(* IEC 61131-3 sources: TwinAxisLab/openplc/cobot-6dof-smart-demo, 8 files *)

(* ---- cobot_6dof_iot_condition_monitoring.st ---- *)
VAR
  Command AT %QW90 : UINT := 0;
  Status AT %QW91 : UINT := 0;
  ActiveStep AT %QW92 : UINT := 0;
  ElapsedMsOut AT %QW93 : UINT := 0;
  AlarmCode AT %QW94 : UINT := 0;
  ConditionState AT %QW95 : UINT := 3;
  SpeedPermille AT %QW96 : UINT := 0;
  ProgramSignature AT %QW97 : UINT := 2101;
  J1Raw AT %QW100 : INT := 0;
  J2Raw AT %QW101 : INT := 0;
  J3Raw AT %QW102 : INT := 0;
  J4Raw AT %QW103 : INT := 0;
  J5Raw AT %QW104 : INT := 0;
  J6Raw AT %QW105 : INT := 0;
  TemperatureCx100 AT %QW120 : INT := 0;
  HumidityRHx100 AT %QW121 : UINT := 0;
  GyroDpsx100 AT %QW122 : UINT := 0;
  SensorAgeMs AT %QW123 : UINT := 65535;
  SensorValid AT %QW124 : UINT := 0;
  SensorSequence AT %QW125 : UINT := 0;
  SensorQualityBits AT %QW126 : UINT := 0;
  SensorPolicy AT %QW127 : UINT := 0;
  CycleTimer : TON;
  MotionIdleTimer : TON;
  TimerEnabled : BOOL := FALSE;
  ResetTimer : BOOL := TRUE;
  ElapsedMs : DINT := 0;
  SegmentStartMs : DINT := 0;
  SegmentDurationMs : DINT := 1;
  P : REAL := 0.0;
  MotionScale : REAL := 1.0;
  TemperatureC : REAL := 0.0;
  HumidityRH : REAL := 0.0;
  GyroDps : REAL := 0.0;
  J1Deg : REAL := 0.0;
  J2Deg : REAL := -35.0;
  J3Deg : REAL := 75.0;
  J4Deg : REAL := 50.0;
  J5Deg : REAL := 0.0;
  J6Deg : REAL := 0.0;
  TargetJ1 : REAL := 0.0;
  TargetJ2 : REAL := -35.0;
  TargetJ3 : REAL := 75.0;
  TargetJ4 : REAL := 50.0;
  TargetJ5 : REAL := 0.0;
  TargetJ6 : REAL := 0.0;
  SegmentStartJ1 : REAL := 0.0;
  SegmentStartJ2 : REAL := -35.0;
  SegmentStartJ3 : REAL := 75.0;
  SegmentStartJ4 : REAL := 50.0;
  SegmentStartJ5 : REAL := 0.0;
  SegmentStartJ6 : REAL := 0.0;
  PreviousStep : UINT := 0;
  PreviousP : REAL := 0.0;
  ProgressDelta : REAL := 0.0;
  MotionPresent : BOOL := FALSE;
  DegToRadScaled : REAL := 174.5329;
END_VAR

ProgramSignature := 2101;

TemperatureC := INT_TO_REAL(TemperatureCx100) / 100.0;
HumidityRH := UINT_TO_REAL(HumidityRHx100) / 100.0;
GyroDps := UINT_TO_REAL(GyroDpsx100) / 100.0;
MotionPresent := GyroDps >= 3.0;
MotionIdleTimer(IN := NOT MotionPresent, PT := T#2s);

ConditionState := 0;
AlarmCode := 0;
MotionScale := 1.0;
SpeedPermille := 1000;

IF (SensorValid = 0) OR ((SensorQualityBits AND 1) = 0) OR (SensorAgeMs > 2500) THEN
  ConditionState := 3;
  AlarmCode := 4;
  MotionScale := 0.0;
  SpeedPermille := 0;
ELSIF ((SensorPolicy = 0) OR (SensorPolicy = 1)) AND ((SensorQualityBits AND 16) = 0) THEN
  ConditionState := 3;
  AlarmCode := 6;
  MotionScale := 0.0;
  SpeedPermille := 0;
ELSIF (TemperatureC >= 55.0) OR (HumidityRH >= 85.0) OR (GyroDps >= 220.0) THEN
  ConditionState := 2;
  MotionScale := 0.0;
  SpeedPermille := 0;
  IF TemperatureC >= 55.0 THEN
    AlarmCode := 1;
  ELSIF HumidityRH >= 85.0 THEN
    AlarmCode := 2;
  ELSE
    AlarmCode := 3;
  END_IF;
ELSIF (TemperatureC >= 45.0) OR (HumidityRH >= 75.0) OR (GyroDps >= 120.0) THEN
  ConditionState := 1;
  MotionScale := 0.55;
  SpeedPermille := 550;
ELSIF (SensorPolicy = 0) AND (NOT MotionPresent) AND (NOT MotionIdleTimer.Q) THEN
  ConditionState := 2;
  AlarmCode := 5;
  MotionScale := 0.0;
  SpeedPermille := 0;
ELSIF (SensorPolicy = 0) AND MotionPresent THEN
  ConditionState := 2;
  AlarmCode := 5;
  MotionScale := 0.0;
  SpeedPermille := 0;
ELSIF (SensorPolicy = 1) AND (NOT MotionPresent) THEN
  ConditionState := 2;
  AlarmCode := 5;
  MotionScale := 0.0;
  SpeedPermille := 0;
END_IF;

IF Command = 2 THEN
  TimerEnabled := FALSE;
  ResetTimer := TRUE;
  Status := 2;
  ActiveStep := 0;
  ElapsedMsOut := 0;
  J1Deg := 0.0;
  J2Deg := -35.0;
  J3Deg := 75.0;
  J4Deg := 50.0;
  J5Deg := 0.0;
  J6Deg := 0.0;
  PreviousStep := 0;
  PreviousP := 0.0;
ELSIF Command = 0 THEN
  TimerEnabled := FALSE;
  ResetTimer := TRUE;
  Status := 0;
  ActiveStep := 0;
  J1Deg := 0.0 + (INT_TO_REAL(J1Raw) / DegToRadScaled);
  J2Deg := -35.0 + (INT_TO_REAL(J2Raw) / DegToRadScaled);
  J3Deg := 75.0 + (INT_TO_REAL(J3Raw) / DegToRadScaled);
  J4Deg := 50.0 + (INT_TO_REAL(J4Raw) / DegToRadScaled);
  J5Deg := 0.0 + (INT_TO_REAL(J5Raw) / DegToRadScaled);
  J6Deg := 0.0 + (INT_TO_REAL(J6Raw) / DegToRadScaled);
  PreviousStep := 0;
  PreviousP := 0.0;
ELSIF ConditionState >= 2 THEN
  TimerEnabled := FALSE;
  ResetTimer := TRUE;
  Status := 3;
  ActiveStep := 0;
  PreviousStep := 0;
  PreviousP := 0.0;
ELSE
  Status := 1;
  IF ResetTimer THEN
    TimerEnabled := FALSE;
    ResetTimer := FALSE;
  ELSE
    TimerEnabled := TRUE;
  END_IF;

  CycleTimer(IN := TimerEnabled, PT := T#10s);
  ElapsedMs := TIME_TO_DINT(CycleTimer.ET);
  IF ElapsedMs > 10000 THEN ElapsedMs := 10000; END_IF;
  ElapsedMsOut := DINT_TO_UINT(ElapsedMs);

  IF ElapsedMs < 1400 THEN
    ActiveStep := 1; SegmentStartMs := 0; SegmentDurationMs := 1400;
  ELSIF ElapsedMs < 2400 THEN
    ActiveStep := 2; SegmentStartMs := 1400; SegmentDurationMs := 1000;
  ELSIF ElapsedMs < 3200 THEN
    ActiveStep := 3; SegmentStartMs := 2400; SegmentDurationMs := 800;
  ELSIF ElapsedMs < 5600 THEN
    ActiveStep := 4; SegmentStartMs := 3200; SegmentDurationMs := 2400;
  ELSIF ElapsedMs < 7600 THEN
    ActiveStep := 5; SegmentStartMs := 5600; SegmentDurationMs := 2000;
  ELSE
    ActiveStep := 6; SegmentStartMs := 7600; SegmentDurationMs := 2400;
  END_IF;

  IF ActiveStep <> PreviousStep THEN
    SegmentStartJ1 := J1Deg;
    SegmentStartJ2 := J2Deg;
    SegmentStartJ3 := J3Deg;
    SegmentStartJ4 := J4Deg;
    SegmentStartJ5 := J5Deg;
    SegmentStartJ6 := J6Deg;
    PreviousStep := ActiveStep;
    PreviousP := 0.0;
  END_IF;

  P := DINT_TO_REAL(ElapsedMs - SegmentStartMs) / DINT_TO_REAL(SegmentDurationMs);
  IF P < 0.0 THEN P := 0.0; END_IF;
  IF P > 1.0 THEN P := 1.0; END_IF;
  P := P * P * (3.0 - (2.0 * P));
  ProgressDelta := P - PreviousP;
  IF ProgressDelta < 0.0 THEN ProgressDelta := 0.0; END_IF;
  IF ProgressDelta > 1.0 THEN ProgressDelta := 1.0; END_IF;
  PreviousP := P;

  IF ActiveStep = 1 THEN
    TargetJ1 := -55.0; TargetJ2 := -10.0; TargetJ3 := 85.0; TargetJ4 := 25.0;
    TargetJ5 := 0.0;
    TargetJ6 := 0.0;
  ELSIF ActiveStep = 2 THEN
    TargetJ1 := -55.0;
    TargetJ2 := 15.0; TargetJ3 := 80.0; TargetJ4 := -5.0;
    TargetJ5 := 0.0;
    TargetJ6 := 0.0;
  ELSIF ActiveStep = 3 THEN
    TargetJ1 := -55.0;
    TargetJ2 := 15.0;
    TargetJ3 := 80.0;
    TargetJ4 := -5.0;
    TargetJ5 := 0.0;
    TargetJ6 := 90.0;
  ELSIF ActiveStep = 4 THEN
    TargetJ1 := 50.0; TargetJ2 := -10.0; TargetJ3 := 85.0; TargetJ4 := 25.0;
    TargetJ5 := 0.0;
    TargetJ6 := 90.0;
  ELSIF ActiveStep = 5 THEN
    TargetJ1 := 50.0;
    TargetJ2 := 15.0; TargetJ3 := 80.0; TargetJ4 := -5.0;
    TargetJ5 := 30.0; TargetJ6 := -90.0;
  ELSE
    TargetJ1 := 0.0; TargetJ2 := -35.0; TargetJ3 := 75.0;
    TargetJ4 := 50.0; TargetJ5 := 0.0; TargetJ6 := 0.0;
  END_IF;

  J1Deg := J1Deg + ((TargetJ1 - SegmentStartJ1) * ProgressDelta * MotionScale);
  J2Deg := J2Deg + ((TargetJ2 - SegmentStartJ2) * ProgressDelta * MotionScale);
  J3Deg := J3Deg + ((TargetJ3 - SegmentStartJ3) * ProgressDelta * MotionScale);
  J4Deg := J4Deg + ((TargetJ4 - SegmentStartJ4) * ProgressDelta * MotionScale);
  J5Deg := J5Deg + ((TargetJ5 - SegmentStartJ5) * ProgressDelta * MotionScale);
  J6Deg := J6Deg + ((TargetJ6 - SegmentStartJ6) * ProgressDelta * MotionScale);

  IF CycleTimer.Q THEN ResetTimer := TRUE; END_IF;
END_IF;

J1Raw := REAL_TO_INT((J1Deg - 0.0) * DegToRadScaled);
J2Raw := REAL_TO_INT((J2Deg - (-35.0)) * DegToRadScaled);
J3Raw := REAL_TO_INT((J3Deg - 75.0) * DegToRadScaled);
J4Raw := REAL_TO_INT((J4Deg - 50.0) * DegToRadScaled);
J5Raw := REAL_TO_INT((J5Deg - 0.0) * DegToRadScaled);
J6Raw := REAL_TO_INT((J6Deg - 0.0) * DegToRadScaled);

(* ---- cobot_6dof_iot_condition_monitoring_old.st ---- *)
  VAR
    Command : UINT AT %QW90 := 0;
    Status : UINT AT %QW91 := 0;
    ActiveStep : UINT AT %QW92 := 0;
    ElapsedMsOut : UINT AT %QW93 := 0;
    AlarmCode : UINT AT %QW94 := 0;
    ConditionState : UINT AT %QW95 := 3;
    SpeedPermille : UINT AT %QW96 := 0;
    ProgramSignature : UINT AT %QW97 := 2101;
    J1Raw : INT AT %QW100 := 0;
    J2Raw : INT AT %QW101 := 0;
    J3Raw : INT AT %QW102 := 0;
    J4Raw : INT AT %QW103 := 0;
    J5Raw : INT AT %QW104 := 0;
    J6Raw : INT AT %QW105 := 0;
    TemperatureCx100 : INT AT %QW120 := 0;
    HumidityRHx100 : UINT AT %QW121 := 0;
    GyroDpsx100 : UINT AT %QW122 := 0;
    SensorAgeMs : UINT AT %QW123 := 65535;
    SensorValid : UINT AT %QW124 := 0;
    SensorSequence : UINT AT %QW125 := 0;
    SensorQualityBits : UINT AT %QW126 := 0;
    SensorPolicy : UINT AT %QW127 := 1;
    CycleTimer : TON;
    MotionIdleTimer : TON;
    TimerEnabled : BOOL := FALSE;
    ResetTimer : BOOL := TRUE;
    ElapsedMs : DINT := 0;
    SegmentStartMs : DINT := 0;
    SegmentDurationMs : DINT := 1;
    P : REAL := 0.0;
    MotionScale : REAL := 1.0;
    TemperatureC : REAL := 0.0;
    HumidityRH : REAL := 0.0;
    GyroDps : REAL := 0.0;
    J1Deg : REAL := 0.0;
    J2Deg : REAL := -35.0;
    J3Deg : REAL := 75.0;
    J4Deg : REAL := 50.0;
    J5Deg : REAL := 0.0;
    J6Deg : REAL := 0.0;
    TargetJ1 : REAL := 0.0;
    TargetJ2 : REAL := -35.0;
    TargetJ3 : REAL := 75.0;
    TargetJ4 : REAL := 50.0;
    TargetJ5 : REAL := 0.0;
    TargetJ6 : REAL := 0.0;
    MotionPresent : BOOL := FALSE;
    DegToRadScaled : REAL := 174.5329;
  END_VAR

TemperatureC := INT_TO_REAL(TemperatureCx100) / 100.0;
HumidityRH := UINT_TO_REAL(HumidityRHx100) / 100.0;
GyroDps := UINT_TO_REAL(GyroDpsx100) / 100.0;
MotionPresent := GyroDps >= 3.0;
MotionIdleTimer(IN := (SensorPolicy = 1) AND (NOT MotionPresent), PT := T#2s);

ConditionState := 0;
AlarmCode := 0;
MotionScale := 1.0;
SpeedPermille := 1000;

IF (SensorValid = 0) OR ((SensorQualityBits AND 1) = 0) OR (SensorAgeMs > 2500) THEN
  ConditionState := 3;
  AlarmCode := 4;
  MotionScale := 0.0;
  SpeedPermille := 0;
ELSIF (SensorPolicy = 1) AND ((SensorQualityBits AND 16) = 0) THEN
  ConditionState := 3;
  AlarmCode := 6;
  MotionScale := 0.0;
  SpeedPermille := 0;
ELSIF (SensorPolicy = 1) AND MotionIdleTimer.Q THEN
  ConditionState := 2;
  AlarmCode := 5;
  MotionScale := 0.0;
  SpeedPermille := 0;
ELSIF (TemperatureC >= 55.0) OR (HumidityRH >= 85.0) OR (GyroDps >= 220.0) THEN
  ConditionState := 2;
  MotionScale := 0.0;
  SpeedPermille := 0;
  IF TemperatureC >= 55.0 THEN
    AlarmCode := 1;
  ELSIF HumidityRH >= 85.0 THEN
    AlarmCode := 2;
  ELSE
    AlarmCode := 3;
  END_IF;
ELSIF (TemperatureC >= 45.0) OR (HumidityRH >= 75.0) OR (GyroDps >= 120.0) THEN
  ConditionState := 1;
  MotionScale := 0.55;
  SpeedPermille := 550;
END_IF;

IF Command = 2 THEN
  TimerEnabled := FALSE;
  ResetTimer := TRUE;
  Status := 2;
  ActiveStep := 0;
  ElapsedMsOut := 0;
  J1Deg := 0.0;
  J2Deg := -35.0;
  J3Deg := 75.0;
  J4Deg := 50.0;
  J5Deg := 0.0;
  J6Deg := 0.0;
ELSIF Command = 0 THEN
  TimerEnabled := FALSE;
  ResetTimer := TRUE;
  Status := 0;
  ActiveStep := 0;
  J1Deg := 0.0 + (INT_TO_REAL(J1Raw) / DegToRadScaled);
  J2Deg := -35.0 + (INT_TO_REAL(J2Raw) / DegToRadScaled);
  J3Deg := 75.0 + (INT_TO_REAL(J3Raw) / DegToRadScaled);
  J4Deg := 50.0 + (INT_TO_REAL(J4Raw) / DegToRadScaled);
  J5Deg := 0.0 + (INT_TO_REAL(J5Raw) / DegToRadScaled);
  J6Deg := 0.0 + (INT_TO_REAL(J6Raw) / DegToRadScaled);
ELSIF ConditionState >= 2 THEN
  TimerEnabled := FALSE;
  ResetTimer := TRUE;
  Status := 3;
  ActiveStep := 0;
ELSE
  Status := 1;
  IF ResetTimer THEN
    TimerEnabled := FALSE;
    ResetTimer := FALSE;
  ELSE
    TimerEnabled := TRUE;
  END_IF;

  CycleTimer(IN := TimerEnabled, PT := T#10s);
  ElapsedMs := TIME_TO_DINT(CycleTimer.ET);
  IF ElapsedMs > 10000 THEN ElapsedMs := 10000; END_IF;
  ElapsedMsOut := DINT_TO_UINT(ElapsedMs);

  IF ElapsedMs < 1400 THEN
    ActiveStep := 1; SegmentStartMs := 0; SegmentDurationMs := 1400;
  ELSIF ElapsedMs < 2400 THEN
    ActiveStep := 2; SegmentStartMs := 1400; SegmentDurationMs := 1000;
  ELSIF ElapsedMs < 3200 THEN
    ActiveStep := 3; SegmentStartMs := 2400; SegmentDurationMs := 800;
  ELSIF ElapsedMs < 5600 THEN
    ActiveStep := 4; SegmentStartMs := 3200; SegmentDurationMs := 2400;
  ELSIF ElapsedMs < 7600 THEN
    ActiveStep := 5; SegmentStartMs := 5600; SegmentDurationMs := 2000;
  ELSE
    ActiveStep := 6; SegmentStartMs := 7600; SegmentDurationMs := 2400;
  END_IF;

  P := DINT_TO_REAL(ElapsedMs - SegmentStartMs) / DINT_TO_REAL(SegmentDurationMs);
  IF P < 0.0 THEN P := 0.0; END_IF;
  IF P > 1.0 THEN P := 1.0; END_IF;
  P := P * P * (3.0 - (2.0 * P));

  IF ActiveStep = 1 THEN
    TargetJ1 := 0.0 + ((-55.0 - 0.0) * P);
    TargetJ2 := -35.0 + ((-10.0 - (-35.0)) * P);
    TargetJ3 := 75.0 + ((85.0 - 75.0) * P);
    TargetJ4 := 50.0 + ((25.0 - 50.0) * P);
    TargetJ5 := 0.0;
    TargetJ6 := 0.0;
  ELSIF ActiveStep = 2 THEN
    TargetJ1 := -55.0;
    TargetJ2 := -10.0 + ((15.0 - (-10.0)) * P);
    TargetJ3 := 85.0 + ((80.0 - 85.0) * P);
    TargetJ4 := 25.0 + ((-5.0 - 25.0) * P);
    TargetJ5 := 0.0;
    TargetJ6 := 0.0;
  ELSIF ActiveStep = 3 THEN
    TargetJ1 := -55.0;
    TargetJ2 := 15.0;
    TargetJ3 := 80.0;
    TargetJ4 := -5.0;
    TargetJ5 := 0.0;
    TargetJ6 := 0.0 + ((90.0 - 0.0) * P);
  ELSIF ActiveStep = 4 THEN
    TargetJ1 := -55.0 + ((50.0 - (-55.0)) * P);
    TargetJ2 := 15.0 + ((-10.0 - 15.0) * P);
    TargetJ3 := 80.0 + ((85.0 - 80.0) * P);
    TargetJ4 := -5.0 + ((25.0 - (-5.0)) * P);
    TargetJ5 := 0.0;
    TargetJ6 := 90.0;
  ELSIF ActiveStep = 5 THEN
    TargetJ1 := 50.0;
    TargetJ2 := -10.0 + ((15.0 - (-10.0)) * P);
    TargetJ3 := 85.0 + ((80.0 - 85.0) * P);
    TargetJ4 := 25.0 + ((-5.0 - 25.0) * P);
    TargetJ5 := 0.0 + ((30.0 - 0.0) * P);
    TargetJ6 := 90.0 + ((-90.0 - 90.0) * P);
  ELSE
    TargetJ1 := 50.0 + ((0.0 - 50.0) * P);
    TargetJ2 := 15.0 + ((-35.0 - 15.0) * P);
    TargetJ3 := 80.0 + ((75.0 - 80.0) * P);
    TargetJ4 := -5.0 + ((50.0 - (-5.0)) * P);
    TargetJ5 := 30.0 + ((0.0 - 30.0) * P);
    TargetJ6 := -90.0 + ((0.0 - (-90.0)) * P);
  END_IF;

  J1Deg := 0.0 + ((TargetJ1 - 0.0) * MotionScale);
  J2Deg := -35.0 + ((TargetJ2 - (-35.0)) * MotionScale);
  J3Deg := 75.0 + ((TargetJ3 - 75.0) * MotionScale);
  J4Deg := 50.0 + ((TargetJ4 - 50.0) * MotionScale);
  J5Deg := 0.0 + ((TargetJ5 - 0.0) * MotionScale);
  J6Deg := 0.0 + ((TargetJ6 - 0.0) * MotionScale);

  IF CycleTimer.Q THEN ResetTimer := TRUE; END_IF;
END_IF;

J1Raw := REAL_TO_INT((J1Deg - 0.0) * DegToRadScaled);
J2Raw := REAL_TO_INT((J2Deg - (-35.0)) * DegToRadScaled);
J3Raw := REAL_TO_INT((J3Deg - 75.0) * DegToRadScaled);
J4Raw := REAL_TO_INT((J4Deg - 50.0) * DegToRadScaled);
J5Raw := REAL_TO_INT((J5Deg - 0.0) * DegToRadScaled);
J6Raw := REAL_TO_INT((J6Deg - 0.0) * DegToRadScaled);

(* ---- cobot_6dof_iot_condition_monitoring_old_07_10_2026.st ---- *)
VAR
  Command AT %QW90 : UINT := 0;
  Status AT %QW91 : UINT := 0;
  ActiveStep AT %QW92 : UINT := 0;
  ElapsedMsOut AT %QW93 : UINT := 0;
  AlarmCode AT %QW94 : UINT := 0;
  ConditionState AT %QW95 : UINT := 3;
  SpeedPermille AT %QW96 : UINT := 0;
  ProgramSignature AT %QW97 : UINT := 2101;
  J1Raw AT %QW100 : INT := 0;
  J2Raw AT %QW101 : INT := 0;
  J3Raw AT %QW102 : INT := 0;
  J4Raw AT %QW103 : INT := 0;
  J5Raw AT %QW104 : INT := 0;
  J6Raw AT %QW105 : INT := 0;
  TemperatureCx100 AT %QW120 : INT := 0;
  HumidityRHx100 AT %QW121 : UINT := 0;
  GyroDpsx100 AT %QW122 : UINT := 0;
  SensorAgeMs AT %QW123 : UINT := 65535;
  SensorValid AT %QW124 : UINT := 0;
  SensorSequence AT %QW125 : UINT := 0;
  SensorQualityBits AT %QW126 : UINT := 0;
  SensorPolicy AT %QW127 : UINT := 1;
  CycleTimer : TON;
  MotionIdleTimer : TON;
  TimerEnabled : BOOL := FALSE;
  ResetTimer : BOOL := TRUE;
  ElapsedMs : DINT := 0;
  SegmentStartMs : DINT := 0;
  SegmentDurationMs : DINT := 1;
  P : REAL := 0.0;
  MotionScale : REAL := 1.0;
  TemperatureC : REAL := 0.0;
  HumidityRH : REAL := 0.0;
  GyroDps : REAL := 0.0;
  J1Deg : REAL := 0.0;
  J2Deg : REAL := -35.0;
  J3Deg : REAL := 75.0;
  J4Deg : REAL := 50.0;
  J5Deg : REAL := 0.0;
  J6Deg : REAL := 0.0;
  TargetJ1 : REAL := 0.0;
  TargetJ2 : REAL := -35.0;
  TargetJ3 : REAL := 75.0;
  TargetJ4 : REAL := 50.0;
  TargetJ5 : REAL := 0.0;
  TargetJ6 : REAL := 0.0;
  SegmentStartJ1 : REAL := 0.0;
  SegmentStartJ2 : REAL := -35.0;
  SegmentStartJ3 : REAL := 75.0;
  SegmentStartJ4 : REAL := 50.0;
  SegmentStartJ5 : REAL := 0.0;
  SegmentStartJ6 : REAL := 0.0;
  PreviousStep : UINT := 0;
  PreviousP : REAL := 0.0;
  ProgressDelta : REAL := 0.0;
  MotionPresent : BOOL := FALSE;
  DegToRadScaled : REAL := 174.5329;
END_VAR

ProgramSignature := 2101;

TemperatureC := INT_TO_REAL(TemperatureCx100) / 100.0;
HumidityRH := UINT_TO_REAL(HumidityRHx100) / 100.0;
GyroDps := UINT_TO_REAL(GyroDpsx100) / 100.0;
MotionPresent := GyroDps >= 3.0;
MotionIdleTimer(IN := (SensorPolicy = 1) AND (NOT MotionPresent), PT := T#2s);

ConditionState := 0;
AlarmCode := 0;
MotionScale := 1.0;
SpeedPermille := 1000;

IF (SensorValid = 0) OR ((SensorQualityBits AND 1) = 0) OR (SensorAgeMs > 2500) THEN
  ConditionState := 3;
  AlarmCode := 4;
  MotionScale := 0.0;
  SpeedPermille := 0;
ELSIF (SensorPolicy = 1) AND ((SensorQualityBits AND 16) = 0) THEN
  ConditionState := 3;
  AlarmCode := 6;
  MotionScale := 0.0;
  SpeedPermille := 0;
ELSIF (SensorPolicy = 1) AND MotionIdleTimer.Q THEN
  ConditionState := 2;
  AlarmCode := 5;
  MotionScale := 0.0;
  SpeedPermille := 0;
ELSIF (TemperatureC >= 55.0) OR (HumidityRH >= 85.0) OR (GyroDps >= 220.0) THEN
  ConditionState := 2;
  MotionScale := 0.0;
  SpeedPermille := 0;
  IF TemperatureC >= 55.0 THEN
    AlarmCode := 1;
  ELSIF HumidityRH >= 85.0 THEN
    AlarmCode := 2;
  ELSE
    AlarmCode := 3;
  END_IF;
ELSIF (TemperatureC >= 45.0) OR (HumidityRH >= 75.0) OR (GyroDps >= 120.0) THEN
  ConditionState := 1;
  MotionScale := 0.55;
  SpeedPermille := 550;
END_IF;

IF Command = 2 THEN
  TimerEnabled := FALSE;
  ResetTimer := TRUE;
  Status := 2;
  ActiveStep := 0;
  ElapsedMsOut := 0;
  J1Deg := 0.0;
  J2Deg := -35.0;
  J3Deg := 75.0;
  J4Deg := 50.0;
  J5Deg := 0.0;
  J6Deg := 0.0;
  PreviousStep := 0;
  PreviousP := 0.0;
ELSIF Command = 0 THEN
  TimerEnabled := FALSE;
  ResetTimer := TRUE;
  Status := 0;
  ActiveStep := 0;
  J1Deg := 0.0 + (INT_TO_REAL(J1Raw) / DegToRadScaled);
  J2Deg := -35.0 + (INT_TO_REAL(J2Raw) / DegToRadScaled);
  J3Deg := 75.0 + (INT_TO_REAL(J3Raw) / DegToRadScaled);
  J4Deg := 50.0 + (INT_TO_REAL(J4Raw) / DegToRadScaled);
  J5Deg := 0.0 + (INT_TO_REAL(J5Raw) / DegToRadScaled);
  J6Deg := 0.0 + (INT_TO_REAL(J6Raw) / DegToRadScaled);
  PreviousStep := 0;
  PreviousP := 0.0;
ELSIF ConditionState >= 2 THEN
  TimerEnabled := FALSE;
  ResetTimer := TRUE;
  Status := 3;
  ActiveStep := 0;
  PreviousStep := 0;
  PreviousP := 0.0;
ELSE
  Status := 1;
  IF ResetTimer THEN
    TimerEnabled := FALSE;
    ResetTimer := FALSE;
  ELSE
    TimerEnabled := TRUE;
  END_IF;

  CycleTimer(IN := TimerEnabled, PT := T#10s);
  ElapsedMs := TIME_TO_DINT(CycleTimer.ET);
  IF ElapsedMs > 10000 THEN ElapsedMs := 10000; END_IF;
  ElapsedMsOut := DINT_TO_UINT(ElapsedMs);

  IF ElapsedMs < 1400 THEN
    ActiveStep := 1; SegmentStartMs := 0; SegmentDurationMs := 1400;
  ELSIF ElapsedMs < 2400 THEN
    ActiveStep := 2; SegmentStartMs := 1400; SegmentDurationMs := 1000;
  ELSIF ElapsedMs < 3200 THEN
    ActiveStep := 3; SegmentStartMs := 2400; SegmentDurationMs := 800;
  ELSIF ElapsedMs < 5600 THEN
    ActiveStep := 4; SegmentStartMs := 3200; SegmentDurationMs := 2400;
  ELSIF ElapsedMs < 7600 THEN
    ActiveStep := 5; SegmentStartMs := 5600; SegmentDurationMs := 2000;
  ELSE
    ActiveStep := 6; SegmentStartMs := 7600; SegmentDurationMs := 2400;
  END_IF;

  IF ActiveStep <> PreviousStep THEN
    SegmentStartJ1 := J1Deg;
    SegmentStartJ2 := J2Deg;
    SegmentStartJ3 := J3Deg;
    SegmentStartJ4 := J4Deg;
    SegmentStartJ5 := J5Deg;
    SegmentStartJ6 := J6Deg;
    PreviousStep := ActiveStep;
    PreviousP := 0.0;
  END_IF;

  P := DINT_TO_REAL(ElapsedMs - SegmentStartMs) / DINT_TO_REAL(SegmentDurationMs);
  IF P < 0.0 THEN P := 0.0; END_IF;
  IF P > 1.0 THEN P := 1.0; END_IF;
  P := P * P * (3.0 - (2.0 * P));
  ProgressDelta := P - PreviousP;
  IF ProgressDelta < 0.0 THEN ProgressDelta := 0.0; END_IF;
  IF ProgressDelta > 1.0 THEN ProgressDelta := 1.0; END_IF;
  PreviousP := P;

  IF ActiveStep = 1 THEN
    TargetJ1 := -55.0; TargetJ2 := -10.0; TargetJ3 := 85.0; TargetJ4 := 25.0;
    TargetJ5 := 0.0;
    TargetJ6 := 0.0;
  ELSIF ActiveStep = 2 THEN
    TargetJ1 := -55.0;
    TargetJ2 := 15.0; TargetJ3 := 80.0; TargetJ4 := -5.0;
    TargetJ5 := 0.0;
    TargetJ6 := 0.0;
  ELSIF ActiveStep = 3 THEN
    TargetJ1 := -55.0;
    TargetJ2 := 15.0;
    TargetJ3 := 80.0;
    TargetJ4 := -5.0;
    TargetJ5 := 0.0;
    TargetJ6 := 90.0;
  ELSIF ActiveStep = 4 THEN
    TargetJ1 := 50.0; TargetJ2 := -10.0; TargetJ3 := 85.0; TargetJ4 := 25.0;
    TargetJ5 := 0.0;
    TargetJ6 := 90.0;
  ELSIF ActiveStep = 5 THEN
    TargetJ1 := 50.0;
    TargetJ2 := 15.0; TargetJ3 := 80.0; TargetJ4 := -5.0;
    TargetJ5 := 30.0; TargetJ6 := -90.0;
  ELSE
    TargetJ1 := 0.0; TargetJ2 := -35.0; TargetJ3 := 75.0;
    TargetJ4 := 50.0; TargetJ5 := 0.0; TargetJ6 := 0.0;
  END_IF;

  J1Deg := J1Deg + ((TargetJ1 - SegmentStartJ1) * ProgressDelta * MotionScale);
  J2Deg := J2Deg + ((TargetJ2 - SegmentStartJ2) * ProgressDelta * MotionScale);
  J3Deg := J3Deg + ((TargetJ3 - SegmentStartJ3) * ProgressDelta * MotionScale);
  J4Deg := J4Deg + ((TargetJ4 - SegmentStartJ4) * ProgressDelta * MotionScale);
  J5Deg := J5Deg + ((TargetJ5 - SegmentStartJ5) * ProgressDelta * MotionScale);
  J6Deg := J6Deg + ((TargetJ6 - SegmentStartJ6) * ProgressDelta * MotionScale);

  IF CycleTimer.Q THEN ResetTimer := TRUE; END_IF;
END_IF;

J1Raw := REAL_TO_INT((J1Deg - 0.0) * DegToRadScaled);
J2Raw := REAL_TO_INT((J2Deg - (-35.0)) * DegToRadScaled);
J3Raw := REAL_TO_INT((J3Deg - 75.0) * DegToRadScaled);
J4Raw := REAL_TO_INT((J4Deg - 50.0) * DegToRadScaled);
J5Raw := REAL_TO_INT((J5Deg - 0.0) * DegToRadScaled);
J6Raw := REAL_TO_INT((J6Deg - 0.0) * DegToRadScaled);

(* ---- cobot_6dof_smart_demo.st ---- *)
VAR
  Command AT %QW90 : UINT := 1;
  Status AT %QW91 : UINT := 1;
  ActiveStep AT %QW92 : UINT := 0;
  ElapsedMsOut AT %QW93 : UINT := 0;
  ProgramSignature AT %QW97 : UINT := 2101;
  J1Raw AT %QW100 : INT := 0;
  J2Raw AT %QW101 : INT := 0;
  J3Raw AT %QW102 : INT := 0;
  J4Raw AT %QW103 : INT := 0;
  J5Raw AT %QW104 : INT := 0;
  J6Raw AT %QW105 : INT := 0;
  CycleTimer : TON;
  TimerEnabled : BOOL := TRUE;
  ResetTimer : BOOL := FALSE;
  ElapsedMs : DINT := 0;
  SegmentStartMs : DINT := 0;
  SegmentDurationMs : DINT := 1;
  P : REAL := 0.0;
  J1Deg : REAL := 0.0;
  J2Deg : REAL := -35.0;
  J3Deg : REAL := 75.0;
  J4Deg : REAL := 50.0;
  J5Deg : REAL := 0.0;
  J6Deg : REAL := 0.0;
  DegToRadScaled : REAL := 174.5329;
END_VAR

ProgramSignature := 2101;

IF Command = 2 THEN
  TimerEnabled := FALSE; Status := 2; ActiveStep := 0; ElapsedMsOut := 0;
  J1Deg := 0.0; J2Deg := -35.0; J3Deg := 75.0;
  J4Deg := 50.0; J5Deg := 0.0; J6Deg := 0.0;
ELSIF Command = 0 THEN
  TimerEnabled := FALSE; Status := 0; ActiveStep := 0;
  J1Deg := 0.0 + (INT_TO_REAL(J1Raw) / DegToRadScaled);
  J2Deg := -35.0 + (INT_TO_REAL(J2Raw) / DegToRadScaled);
  J3Deg := 75.0 + (INT_TO_REAL(J3Raw) / DegToRadScaled);
  J4Deg := 50.0 + (INT_TO_REAL(J4Raw) / DegToRadScaled);
  J5Deg := 0.0 + (INT_TO_REAL(J5Raw) / DegToRadScaled);
  J6Deg := 0.0 + (INT_TO_REAL(J6Raw) / DegToRadScaled);
ELSE
  Status := 1;
  IF ResetTimer THEN
    TimerEnabled := FALSE; ResetTimer := FALSE;
  ELSE
    TimerEnabled := TRUE;
  END_IF;

  CycleTimer(IN := TimerEnabled, PT := T#10s);
  ElapsedMs := TIME_TO_DINT(CycleTimer.ET);
  IF ElapsedMs > 10000 THEN ElapsedMs := 10000; END_IF;
  ElapsedMsOut := DINT_TO_UINT(ElapsedMs);

  IF ElapsedMs < 1400 THEN
    ActiveStep := 1; SegmentStartMs := 0; SegmentDurationMs := 1400;
  ELSIF ElapsedMs < 2400 THEN
    ActiveStep := 2; SegmentStartMs := 1400; SegmentDurationMs := 1000;
  ELSIF ElapsedMs < 3200 THEN
    ActiveStep := 3; SegmentStartMs := 2400; SegmentDurationMs := 800;
  ELSIF ElapsedMs < 5600 THEN
    ActiveStep := 4; SegmentStartMs := 3200; SegmentDurationMs := 2400;
  ELSIF ElapsedMs < 7600 THEN
    ActiveStep := 5; SegmentStartMs := 5600; SegmentDurationMs := 2000;
  ELSE
    ActiveStep := 6; SegmentStartMs := 7600; SegmentDurationMs := 2400;
  END_IF;

  IF SegmentDurationMs > 0 THEN
    P := DINT_TO_REAL(ElapsedMs - SegmentStartMs) / DINT_TO_REAL(SegmentDurationMs);
    IF P < 0.0 THEN P := 0.0; ELSIF P > 1.0 THEN P := 1.0; END_IF;
    P := P * P * (3.0 - (2.0 * P));
  ELSE
    P := 0.0;
  END_IF;

  IF ActiveStep = 1 THEN
    J1Deg := 0.0 + ((-55.0 - 0.0) * P);
    J2Deg := -35.0 + ((-10.0 - (-35.0)) * P);
    J3Deg := 75.0 + ((85.0 - 75.0) * P);
    J4Deg := 50.0 + ((25.0 - 50.0) * P);
    J5Deg := 0.0;
    J6Deg := 0.0;
  ELSIF ActiveStep = 2 THEN
    J1Deg := -55.0;
    J2Deg := -10.0 + ((15.0 - (-10.0)) * P);
    J3Deg := 85.0 + ((80.0 - 85.0) * P);
    J4Deg := 25.0 + ((-5.0 - 25.0) * P);
    J5Deg := 0.0;
    J6Deg := 0.0;
  ELSIF ActiveStep = 3 THEN
    J1Deg := -55.0;
    J2Deg := 15.0;
    J3Deg := 80.0;
    J4Deg := -5.0;
    J5Deg := 0.0;
    J6Deg := 0.0 + ((90.0 - 0.0) * P);
  ELSIF ActiveStep = 4 THEN
    J1Deg := -55.0 + ((50.0 - (-55.0)) * P);
    J2Deg := 15.0 + ((-10.0 - 15.0) * P);
    J3Deg := 80.0 + ((85.0 - 80.0) * P);
    J4Deg := -5.0 + ((25.0 - (-5.0)) * P);
    J5Deg := 0.0;
    J6Deg := 90.0;
  ELSIF ActiveStep = 5 THEN
    J1Deg := 50.0;
    J2Deg := -10.0 + ((15.0 - (-10.0)) * P);
    J3Deg := 85.0 + ((80.0 - 85.0) * P);
    J4Deg := 25.0 + ((-5.0 - 25.0) * P);
    J5Deg := 0.0 + ((30.0 - 0.0) * P);
    J6Deg := 90.0 + ((-90.0 - 90.0) * P);
  ELSE
    J1Deg := 50.0 + ((0.0 - 50.0) * P);
    J2Deg := 15.0 + ((-35.0 - 15.0) * P);
    J3Deg := 80.0 + ((75.0 - 80.0) * P);
    J4Deg := -5.0 + ((50.0 - (-5.0)) * P);
    J5Deg := 30.0 + ((0.0 - 30.0) * P);
    J6Deg := -90.0 + ((0.0 - (-90.0)) * P);
  END_IF;

  IF CycleTimer.Q THEN ResetTimer := TRUE; END_IF;
END_IF;

J1Raw := REAL_TO_INT((J1Deg - 0.0) * DegToRadScaled);
J2Raw := REAL_TO_INT((J2Deg - (-35.0)) * DegToRadScaled);
J3Raw := REAL_TO_INT((J3Deg - 75.0) * DegToRadScaled);
J4Raw := REAL_TO_INT((J4Deg - 50.0) * DegToRadScaled);
J5Raw := REAL_TO_INT((J5Deg - 0.0) * DegToRadScaled);
J6Raw := REAL_TO_INT((J6Deg - 0.0) * DegToRadScaled);

(* ---- cobot_6dof_smart_demo_amplified.st ---- *)
VAR
  Command AT %QW90 : UINT := 0;
  Status AT %QW91 : UINT := 0;
  ActiveStep AT %QW92 : UINT := 0;
  ElapsedMsOut AT %QW93 : UINT := 0;
  J1Raw AT %QW100 : INT := 0;
  J2Raw AT %QW101 : INT := -6109;
  J3Raw AT %QW102 : INT := 13090;
  J4Raw AT %QW103 : INT := 8727;
  J5Raw AT %QW104 : INT := 0;
  J6Raw AT %QW105 : INT := 0;
  CycleTimer : TON;
  TimerEnabled : BOOL := FALSE;
  ResetTimer : BOOL := FALSE;
  ElapsedMs : DINT := 0;
  SegmentStartMs : DINT := 0;
  SegmentDurationMs : DINT := 1;
  P : REAL := 0.0;
  J1Deg : REAL := 0.0;
  J2Deg : REAL := -35.0;
  J3Deg : REAL := 75.0;
  J4Deg : REAL := 50.0;
  J5Deg : REAL := 0.0;
  J6Deg : REAL := 0.0;
  DegToRadScaled : REAL := 174.5329;
END_VAR

IF Command = 2 THEN
  TimerEnabled := FALSE;
  ResetTimer := TRUE;
  Status := 2;
  ActiveStep := 0;
  ElapsedMsOut := 0;
  J1Deg := 0.0;
  J2Deg := -35.0;
  J3Deg := 75.0;
  J4Deg := 50.0;
  J5Deg := 0.0;
  J6Deg := 0.0;
ELSIF Command = 0 THEN
  TimerEnabled := FALSE;
  ResetTimer := TRUE;
  Status := 0;
  ActiveStep := 0;
  ElapsedMsOut := 0;
  J1Deg := INT_TO_REAL(J1Raw) / DegToRadScaled;
  J2Deg := INT_TO_REAL(J2Raw) / DegToRadScaled;
  J3Deg := INT_TO_REAL(J3Raw) / DegToRadScaled;
  J4Deg := INT_TO_REAL(J4Raw) / DegToRadScaled;
  J5Deg := INT_TO_REAL(J5Raw) / DegToRadScaled;
  J6Deg := INT_TO_REAL(J6Raw) / DegToRadScaled;
ELSE
  Status := 1;

  IF ResetTimer THEN
    TimerEnabled := FALSE;
    ResetTimer := FALSE;
  ELSE
    TimerEnabled := TRUE;
  END_IF;

  CycleTimer(IN := TimerEnabled, PT := T#18s);
  ElapsedMs := TIME_TO_DINT(CycleTimer.ET);
  IF ElapsedMs > 18000 THEN ElapsedMs := 18000; END_IF;
  ElapsedMsOut := DINT_TO_UINT(ElapsedMs);

  IF ElapsedMs < 3000 THEN
    ActiveStep := 1;
    SegmentStartMs := 0;
    SegmentDurationMs := 3000;
  ELSIF ElapsedMs < 6000 THEN
    ActiveStep := 2;
    SegmentStartMs := 3000;
    SegmentDurationMs := 3000;
  ELSIF ElapsedMs < 9000 THEN
    ActiveStep := 3;
    SegmentStartMs := 6000;
    SegmentDurationMs := 3000;
  ELSIF ElapsedMs < 12000 THEN
    ActiveStep := 4;
    SegmentStartMs := 9000;
    SegmentDurationMs := 3000;
  ELSIF ElapsedMs < 15000 THEN
    ActiveStep := 5;
    SegmentStartMs := 12000;
    SegmentDurationMs := 3000;
  ELSE
    ActiveStep := 6;
    SegmentStartMs := 15000;
    SegmentDurationMs := 3000;
  END_IF;

  P := DINT_TO_REAL(ElapsedMs - SegmentStartMs) / DINT_TO_REAL(SegmentDurationMs);
  IF P < 0.0 THEN P := 0.0; END_IF;
  IF P > 1.0 THEN P := 1.0; END_IF;
  P := P * P * (3.0 - (2.0 * P));

  IF ActiveStep = 1 THEN
    J1Deg := 0.0 + ((-150.0 - 0.0) * P);
    J2Deg := -35.0 + ((-75.0 - (-35.0)) * P);
    J3Deg := 75.0 + ((110.0 - 75.0) * P);
    J4Deg := 50.0 + ((-90.0 - 50.0) * P);
    J5Deg := 0.0 + ((-80.0 - 0.0) * P);
    J6Deg := 0.0 + ((-160.0 - 0.0) * P);
  ELSIF ActiveStep = 2 THEN
    J1Deg := -150.0;
    J2Deg := -75.0 + ((70.0 - (-75.0)) * P);
    J3Deg := 110.0 + ((145.0 - 110.0) * P);
    J4Deg := -90.0 + ((120.0 - (-90.0)) * P);
    J5Deg := -80.0 + ((100.0 - (-80.0)) * P);
    J6Deg := -160.0 + ((160.0 - (-160.0)) * P);
  ELSIF ActiveStep = 3 THEN
    J1Deg := -150.0 + ((150.0 - (-150.0)) * P);
    J2Deg := 70.0 + ((20.0 - 70.0) * P);
    J3Deg := 145.0 + ((40.0 - 145.0) * P);
    J4Deg := 120.0 + ((-130.0 - 120.0) * P);
    J5Deg := 100.0 + ((-110.0 - 100.0) * P);
    J6Deg := 160.0 + ((-170.0 - 160.0) * P);
  ELSIF ActiveStep = 4 THEN
    J1Deg := 150.0;
    J2Deg := 20.0 + ((-100.0 - 20.0) * P);
    J3Deg := 40.0 + ((130.0 - 40.0) * P);
    J4Deg := -130.0 + ((140.0 - (-130.0)) * P);
    J5Deg := -110.0 + ((120.0 - (-110.0)) * P);
    J6Deg := -170.0 + ((170.0 - (-170.0)) * P);
  ELSIF ActiveStep = 5 THEN
    J1Deg := 150.0 + ((-110.0 - 150.0) * P);
    J2Deg := -100.0 + ((80.0 - (-100.0)) * P);
    J3Deg := 130.0 + ((25.0 - 130.0) * P);
    J4Deg := 140.0 + ((-140.0 - 140.0) * P);
    J5Deg := 120.0 + ((-120.0 - 120.0) * P);
    J6Deg := 170.0 + ((-165.0 - 170.0) * P);
  ELSE
    J1Deg := -110.0 + ((0.0 - (-110.0)) * P);
    J2Deg := 80.0 + ((-35.0 - 80.0) * P);
    J3Deg := 25.0 + ((75.0 - 25.0) * P);
    J4Deg := -140.0 + ((50.0 - (-140.0)) * P);
    J5Deg := -120.0 + ((0.0 - (-120.0)) * P);
    J6Deg := -165.0 + ((0.0 - (-165.0)) * P);
  END_IF;

  IF CycleTimer.Q THEN ResetTimer := TRUE; END_IF;
END_IF;

IF J1Deg < -170.0 THEN J1Deg := -170.0; END_IF;
IF J1Deg > 170.0 THEN J1Deg := 170.0; END_IF;
IF J2Deg < -120.0 THEN J2Deg := -120.0; END_IF;
IF J2Deg > 120.0 THEN J2Deg := 120.0; END_IF;
IF J3Deg < -170.0 THEN J3Deg := -170.0; END_IF;
IF J3Deg > 170.0 THEN J3Deg := 170.0; END_IF;
IF J4Deg < -170.0 THEN J4Deg := -170.0; END_IF;
IF J4Deg > 170.0 THEN J4Deg := 170.0; END_IF;
IF J5Deg < -170.0 THEN J5Deg := -170.0; END_IF;
IF J5Deg > 170.0 THEN J5Deg := 170.0; END_IF;
IF J6Deg < -175.0 THEN J6Deg := -175.0; END_IF;
IF J6Deg > 175.0 THEN J6Deg := 175.0; END_IF;

J1Raw := REAL_TO_INT(J1Deg * DegToRadScaled);
J2Raw := REAL_TO_INT(J2Deg * DegToRadScaled);
J3Raw := REAL_TO_INT(J3Deg * DegToRadScaled);
J4Raw := REAL_TO_INT(J4Deg * DegToRadScaled);
J5Raw := REAL_TO_INT(J5Deg * DegToRadScaled);
J6Raw := REAL_TO_INT(J6Deg * DegToRadScaled);

(* ---- cobot_6dof_smart_demo_rectificado.st ---- *)
VAR
  Command AT %QW90 : UINT := 1;
  Status AT %QW91 : UINT := 1;
  ActiveStep AT %QW92 : UINT := 0;
  ElapsedMsOut AT %QW93 : UINT := 0;
  J1Raw AT %QW100 : INT := 0;
  J2Raw AT %QW101 : INT := -6109;
  J3Raw AT %QW102 : INT := 13090;
  J4Raw AT %QW103 : INT := 8727;
  J5Raw AT %QW104 : INT := 0;
  J6Raw AT %QW105 : INT := 0;
  CycleTimer : TON;
  TimerEnabled : BOOL := TRUE;
  ResetTimer : BOOL := FALSE;
  ElapsedMs : DINT := 0;
  SegmentStartMs : DINT := 0;
  SegmentDurationMs : DINT := 1;
  P : REAL := 0.0;
  J1Deg : REAL := 0.0;
  J2Deg : REAL := -35.0;
  J3Deg : REAL := 75.0;
  J4Deg : REAL := 50.0;
  J5Deg : REAL := 0.0;
  J6Deg : REAL := 0.0;
  DegToRadScaled : REAL := 174.5329;
END_VAR

IF Command = 2 THEN
  TimerEnabled := FALSE; Status := 2; ActiveStep := 0; ElapsedMsOut := 0;
  J1Deg := 0.0; J2Deg := -35.0; J3Deg := 75.0;
  J4Deg := 50.0; J5Deg := 0.0; J6Deg := 0.0;
ELSIF Command = 0 THEN
  TimerEnabled := FALSE; Status := 0; ActiveStep := 0;
  J1Deg := INT_TO_REAL(J1Raw) / DegToRadScaled;
  J2Deg := INT_TO_REAL(J2Raw) / DegToRadScaled;
  J3Deg := INT_TO_REAL(J3Raw) / DegToRadScaled;
  J4Deg := INT_TO_REAL(J4Raw) / DegToRadScaled;
  J5Deg := INT_TO_REAL(J5Raw) / DegToRadScaled;
  J6Deg := INT_TO_REAL(J6Raw) / DegToRadScaled;
ELSE
  Status := 1;
  IF ResetTimer THEN
    TimerEnabled := FALSE; ResetTimer := FALSE;
  ELSE
    TimerEnabled := TRUE;
  END_IF;

  CycleTimer(IN := TimerEnabled, PT := T#10s);
  ElapsedMs := TIME_TO_DINT(CycleTimer.ET);
  IF ElapsedMs > 10000 THEN ElapsedMs := 10000; END_IF;
  ElapsedMsOut := DINT_TO_UINT(ElapsedMs);

  IF ElapsedMs < 1400 THEN
    ActiveStep := 1; SegmentStartMs := 0; SegmentDurationMs := 1400;
  ELSIF ElapsedMs < 2400 THEN
    ActiveStep := 2; SegmentStartMs := 1400; SegmentDurationMs := 1000;
  ELSIF ElapsedMs < 3200 THEN
    ActiveStep := 3; SegmentStartMs := 2400; SegmentDurationMs := 800;
  ELSIF ElapsedMs < 5600 THEN
    ActiveStep := 4; SegmentStartMs := 3200; SegmentDurationMs := 2400;
  ELSIF ElapsedMs < 7600 THEN
    ActiveStep := 5; SegmentStartMs := 5600; SegmentDurationMs := 2000;
  ELSE
    ActiveStep := 6; SegmentStartMs := 7600; SegmentDurationMs := 2400;
  END_IF;

  IF SegmentDurationMs > 0 THEN
    P := DINT_TO_REAL(ElapsedMs - SegmentStartMs) / DINT_TO_REAL(SegmentDurationMs);
    IF P < 0.0 THEN P := 0.0; ELSIF P > 1.0 THEN P := 1.0; END_IF;
  ELSE
    P := 0.0;
  END_IF;

  IF ActiveStep = 1 THEN
    J1Deg := 0.0 + ((-55.0 - 0.0) * P);
    J2Deg := -35.0 + ((-10.0 - (-35.0)) * P);
    J3Deg := 75.0 + ((85.0 - 75.0) * P);
    J4Deg := 50.0 + ((25.0 - 50.0) * P);
    J5Deg := 0.0;
    J6Deg := 0.0;
  ELSIF ActiveStep = 2 THEN
    J1Deg := -55.0;
    J2Deg := -10.0 + ((15.0 - (-10.0)) * P);
    J3Deg := 85.0 + ((80.0 - 85.0) * P);
    J4Deg := 25.0 + ((-5.0 - 25.0) * P);
    J5Deg := 0.0;
    J6Deg := 0.0;
  ELSIF ActiveStep = 3 THEN
    J1Deg := -55.0;
    J2Deg := 15.0;
    J3Deg := 80.0;
    J4Deg := -5.0;
    J5Deg := 0.0;
    J6Deg := 0.0 + ((90.0 - 0.0) * P);
  ELSIF ActiveStep = 4 THEN
    J1Deg := -55.0 + ((50.0 - (-55.0)) * P);
    J2Deg := 15.0 + ((-10.0 - 15.0) * P);
    J3Deg := 80.0 + ((85.0 - 80.0) * P);
    J4Deg := -5.0 + ((25.0 - (-5.0)) * P);
    J5Deg := 0.0;
    J6Deg := 90.0;
  ELSIF ActiveStep = 5 THEN
    J1Deg := 50.0;
    J2Deg := -10.0 + ((15.0 - (-10.0)) * P);
    J3Deg := 85.0 + ((80.0 - 85.0) * P);
    J4Deg := 25.0 + ((-5.0 - 25.0) * P);
    J5Deg := 0.0 + ((30.0 - 0.0) * P);
    J6Deg := 90.0 + ((-90.0 - 90.0) * P);
  ELSE
    J1Deg := 50.0 + ((0.0 - 50.0) * P);
    J2Deg := 15.0 + ((-35.0 - 15.0) * P);
    J3Deg := 80.0 + ((75.0 - 80.0) * P);
    J4Deg := -5.0 + ((50.0 - (-5.0)) * P);
    J5Deg := 30.0 + ((0.0 - 30.0) * P);
    J6Deg := -90.0 + ((0.0 - (-90.0)) * P);
  END_IF;

  IF CycleTimer.Q THEN ResetTimer := TRUE; END_IF;
END_IF;

J1Raw := REAL_TO_INT(J1Deg * DegToRadScaled);
J2Raw := REAL_TO_INT(J2Deg * DegToRadScaled);
J3Raw := REAL_TO_INT(J3Deg * DegToRadScaled);
J4Raw := REAL_TO_INT(J4Deg * DegToRadScaled);
J5Raw := REAL_TO_INT(J5Deg * DegToRadScaled);
J6Raw := REAL_TO_INT(J6Deg * DegToRadScaled);

(* ---- FB_FT511938_openplc.st ---- *)
VAR
  Cmd AT %QW0 : UINT := 0;
  Enable AT %QW1 : UINT := 1;
  JogAxis AT %QW2 : INT := 0;
  JogDirection AT %QW3 : INT := 0;
  JogEnable AT %QW4 : UINT := 0;
  HeartbeatSequence AT %QW5 : UINT := 0;

  ManualTarget1High AT %QW6 : UINT := 0;
  ManualTarget1Low AT %QW7 : UINT := 0;
  ManualTarget2High AT %QW8 : UINT := 17302;
  ManualTarget2Low AT %QW9 : UINT := 0;
  ManualTarget3High AT %QW10 : UINT := 17008;
  ManualTarget3Low AT %QW11 : UINT := 0;
  ManualTarget4High AT %QW12 : UINT := 16968;
  ManualTarget4Low AT %QW13 : UINT := 0;

  SensorPolicy AT %QW14 : UINT := 0;
  SensorValid AT %QW15 : UINT := 1;
  SensorQualityBits AT %QW16 : UINT := 17;
  SensorAgeMs AT %QW17 : UINT := 0;
  TemperatureCx100 AT %QW18 : INT := 2200;
  HumidityRHx100 AT %QW19 : UINT := 5000;
  GyroDpsx100 AT %QW20 : UINT := 0;

  SafetyOK AT %QW21 : UINT := 0;
  DrivesReady AT %QW22 : UINT := 0;
  CommFresh AT %QW23 : UINT := 1;
  SensorOK AT %QW24 : UINT := 1;
  HomedMask AT %QW25 : UINT := 15;
  MinLimitMask AT %QW26 : UINT := 0;
  MaxLimitMask AT %QW27 : UINT := 0;
  WiringVerified AT %QW28 : UINT := 0;
  PhysicalOutputEnable AT %QW29 : UINT := 0;

  Pos1High AT %QW30 : UINT := 0;
  Pos1Low AT %QW31 : UINT := 0;
  Pos2High AT %QW32 : UINT := 0;
  Pos2Low AT %QW33 : UINT := 0;
  Pos3High AT %QW34 : UINT := 0;
  Pos3Low AT %QW35 : UINT := 0;
  Pos4High AT %QW36 : UINT := 0;
  Pos4Low AT %QW37 : UINT := 0;
  Target1High AT %QW38 : UINT := 0;
  Target1Low AT %QW39 : UINT := 0;
  Target2High AT %QW40 : UINT := 0;
  Target2Low AT %QW41 : UINT := 0;
  Target3High AT %QW42 : UINT := 0;
  Target3Low AT %QW43 : UINT := 0;
  Target4High AT %QW44 : UINT := 0;
  Target4Low AT %QW45 : UINT := 0;

  Status AT %QW46 : UINT := 0;
  ActiveMode AT %QW47 : UINT := 0;
  ActiveStep AT %QW48 : UINT := 0;
  AlarmCode AT %QW49 : UINT := 0;
  Done AT %QW50 : UINT := 0;
  IoTAlarmCode AT %QW51 : UINT := 0;
  ConditionState AT %QW52 : UINT := 0;
  SpeedPermille AT %QW53 : UINT := 1000;
  CmdQ1toQ8Mask AT %QW54 : UINT := 0;
  RunMask AT %QW55 : UINT := 0;
  DirectionMask AT %QW56 : UINT := 0;
  HeartbeatEcho AT %QW57 : UINT := 0;
  SimulationMode AT %QW58 : UINT := 1;
  StartupReady AT %QW59 : UINT := 0;
  DoneCounter AT %QW60 : UINT := 0;

  SegmentTimer : TON;
  AutoSegmentTimerA : TON;
  AutoSegmentTimerB : TON;
  JogPulseTimer : TON;
  SettleTimer : TON;
  MotionIdleTimer : TON;

  ModeState : UINT := 0;
  LastCmd : UINT := 0;
  Step : UINT := 0;
  ActiveAxis : UINT := 0;
  LastActiveAxis : UINT := 0;
  Fault : UINT := 0;
  SegmentDurationMs : DINT := 1800;
  P : REAL := 0.0;
  SegmentRunning : BOOL := FALSE;
  AutoSegmentReady : BOOL := FALSE;
  AutoSegmentRunning : BOOL := FALSE;
  AutoSegmentDone : BOOL := FALSE;
  AtTarget : BOOL := FALSE;
  AnyMoving : BOOL := FALSE;
  DonePulse : BOOL := FALSE;
  IoTBlock : BOOL := FALSE;
  IoTDegraded : BOOL := FALSE;
  PhysicalPermitted : BOOL := FALSE;
  ManualPermitted : BOOL := FALSE;
  AutoPermitted : BOOL := FALSE;
  AutoMotionAllowed : BOOL := FALSE;
  Permitted : BOOL := FALSE;
  MotionPresent : BOOL := FALSE;
  TemperatureC : REAL := 0.0;
  HumidityRH : REAL := 0.0;
  GyroDps : REAL := 0.0;
  MotionScale : REAL := 1.0;

  Current1 : REAL := 0.0;
  Current2 : REAL := 300.0;
  Current3 : REAL := 60.0;
  Current4 : REAL := 50.0;
  Captured1 : REAL := 0.0;
  Captured2 : REAL := 300.0;
  Captured3 : REAL := 60.0;
  Captured4 : REAL := 50.0;
  SegmentStart1 : REAL := 0.0;
  SegmentStart2 : REAL := 300.0;
  SegmentStart3 : REAL := 60.0;
  SegmentStart4 : REAL := 50.0;
  AutoSegmentStart1 : REAL := 0.0;
  AutoSegmentStart2 : REAL := 300.0;
  AutoSegmentStart3 : REAL := 60.0;
  AutoSegmentStart4 : REAL := 50.0;
  TargetValue : REAL := 0.0;
  ManualValid : BOOL := FALSE;
  DemoTarget1 : REAL := 0.0;
  DemoTarget2 : REAL := 300.0;
  DemoTarget3 : REAL := 60.0;
  DemoTarget4 : REAL := 50.0;
  AxisTarget2 : REAL := 300.0;
  ManualSafeHeight : BOOL := FALSE;
  ManualPhase : UINT := 0;
  ManualPlanActive : BOOL := FALSE;
  ManualRequiresSafeHeight : BOOL := FALSE;
  ManualTargetChanged : BOOL := FALSE;
  ManualAxisTarget2 : REAL := 300.0;
  ManualComplete : BOOL := FALSE;
  ManualTargetError : BOOL := FALSE;
  ManualBaseReady : BOOL := FALSE;
  ManualExtensionReady : BOOL := FALSE;
  ManualSafeHeightReady : BOOL := FALSE;
  ManualHeightReady : BOOL := FALSE;
  ManualGripperReady : BOOL := FALSE;
  StartupDefaultsApplied : BOOL := FALSE;
  RealBits : POINTER TO DWORD;
  RawReal : DWORD := 0;
  RawRealPointer : POINTER TO REAL;
  ManualTarget1 : REAL := 0.0;
  ManualTarget2 : REAL := 300.0;
  ManualTarget3 : REAL := 60.0;
  ManualTarget4 : REAL := 50.0;
  Pos1 : REAL := 0.0;
  Pos2 : REAL := 300.0;
  Pos3 : REAL := 60.0;
  Pos4 : REAL := 50.0;
  Target1 : REAL := 0.0;
  Target2 : REAL := 300.0;
  Target3 : REAL := 60.0;
  Target4 : REAL := 50.0;
END_VAR

IF NOT StartupDefaultsApplied THEN
  IF ((Pos4High = 0) AND (Pos4Low = 0))
     OR (Pos2 < 128.0) OR (Pos2 > 362.0)
     OR (Pos4 < 10.0) OR (Pos4 > 72.0) THEN
    Enable := 1;
    HomedMask := 15;
    SimulationMode := 1;
    Current1 := 0.0;
    Current2 := 300.0;
    Current3 := 60.0;
    Current4 := 50.0;
    Captured1 := 0.0;
    Captured2 := 300.0;
    Captured3 := 60.0;
    Captured4 := 50.0;
    DemoTarget1 := 0.0;
    DemoTarget2 := 300.0;
    DemoTarget3 := 60.0;
    DemoTarget4 := 50.0;
    AxisTarget2 := 300.0;
    ManualAxisTarget2 := 300.0;
  END_IF;
  StartupDefaultsApplied := TRUE;
END_IF;

RawReal := SHL(TO_DWORD(ManualTarget1High), 16) OR TO_DWORD(ManualTarget1Low);
RawRealPointer := ADR(RawReal);
ManualTarget1 := RawRealPointer^;
RawReal := SHL(TO_DWORD(ManualTarget2High), 16) OR TO_DWORD(ManualTarget2Low);
RawRealPointer := ADR(RawReal);
ManualTarget2 := RawRealPointer^;
RawReal := SHL(TO_DWORD(ManualTarget3High), 16) OR TO_DWORD(ManualTarget3Low);
RawRealPointer := ADR(RawReal);
ManualTarget3 := RawRealPointer^;
RawReal := SHL(TO_DWORD(ManualTarget4High), 16) OR TO_DWORD(ManualTarget4Low);
RawRealPointer := ADR(RawReal);
ManualTarget4 := RawRealPointer^;

StartupReady := 1;

HeartbeatEcho := HeartbeatSequence;
TemperatureC := INT_TO_REAL(TemperatureCx100) / 100.0;
HumidityRH := UINT_TO_REAL(HumidityRHx100) / 100.0;
GyroDps := UINT_TO_REAL(GyroDpsx100) / 100.0;
MotionPresent := GyroDps >= 3.0;
MotionIdleTimer(IN := NOT MotionPresent, PT := T#2s);

ConditionState := 0;
IoTAlarmCode := 0;
SpeedPermille := 1000;
MotionScale := 1.0;
IF (SensorValid = 0) OR ((SensorQualityBits AND 1) = 0) OR (SensorAgeMs > 2500) THEN
  ConditionState := 3;
  IoTAlarmCode := 4;
  MotionScale := 0.0;
  SpeedPermille := 0;
ELSIF ((SensorPolicy = 0) OR (SensorPolicy = 1)) AND ((SensorQualityBits AND 16) = 0) THEN
  ConditionState := 3;
  IoTAlarmCode := 6;
  MotionScale := 0.0;
  SpeedPermille := 0;
ELSIF (TemperatureC >= 55.0) OR (HumidityRH >= 85.0) OR (GyroDps >= 220.0) THEN
  ConditionState := 2;
  MotionScale := 0.0;
  SpeedPermille := 0;
  IF TemperatureC >= 55.0 THEN
    IoTAlarmCode := 1;
  ELSIF HumidityRH >= 85.0 THEN
    IoTAlarmCode := 2;
  ELSE
    IoTAlarmCode := 3;
  END_IF;
ELSIF (TemperatureC >= 45.0) OR (HumidityRH >= 75.0) OR (GyroDps >= 120.0) THEN
  ConditionState := 1;
  MotionScale := 0.0;
  SpeedPermille := 550;
ELSIF (SensorPolicy = 0) AND (NOT MotionPresent) AND (NOT MotionIdleTimer.Q) THEN
  ConditionState := 2;
  IoTAlarmCode := 5;
  MotionScale := 0.0;
  SpeedPermille := 0;
ELSIF (SensorPolicy = 0) AND MotionPresent THEN
  ConditionState := 2;
  IoTAlarmCode := 5;
  MotionScale := 0.0;
  SpeedPermille := 0;
ELSIF (SensorPolicy = 1) AND NOT MotionPresent THEN
  ConditionState := 2;
  IoTAlarmCode := 5;
  MotionScale := 0.0;
  SpeedPermille := 0;
END_IF;

IoTBlock := ConditionState >= 2;
IoTDegraded := ConditionState = 1;
PhysicalPermitted := (Enable <> 0) AND (HomedMask = 15)
                     AND ((SimulationMode <> 0)
                          OR ((SafetyOK <> 0) AND (DrivesReady <> 0)
                              AND (WiringVerified <> 0) AND (PhysicalOutputEnable <> 0)));

ManualPermitted := PhysicalPermitted;

AutoMotionAllowed := FALSE;
IF SensorPolicy = 0 THEN
  AutoMotionAllowed := (NOT MotionPresent) AND MotionIdleTimer.Q;
ELSIF SensorPolicy = 1 THEN
  AutoMotionAllowed := MotionPresent;
END_IF;

AutoPermitted := PhysicalPermitted
                 AND (CommFresh <> 0)
                 AND (SensorOK <> 0)
                 AND (SensorValid <> 0)
                 AND ((SensorQualityBits AND 1) <> 0)
                 AND ((SensorQualityBits AND 16) <> 0)
                 AND (SensorAgeMs <= 2500)
                 AND (NOT IoTBlock)
                 AND (NOT IoTDegraded)
                 AND AutoMotionAllowed;

IF ModeState = 1 THEN
  Permitted := AutoPermitted;
ELSE
  Permitted := ManualPermitted;
END_IF;

Pos1 := Current1;
Pos2 := Current2;
Pos3 := Current3;
Pos4 := Current4;

Done := 0;
DonePulse := FALSE;
AnyMoving := FALSE;
AtTarget := FALSE;
ActiveAxis := 0;
Fault := 0;

IF Cmd = 2 THEN
  IF LastCmd <> 2 THEN
    ModeState := 2;
    Step := 0;
    Captured1 := 0.0;
    Captured2 := 300.0;
    Captured3 := 60.0;
    Captured4 := 50.0;
    ManualSafeHeight := FALSE;
    ManualPhase := 0;
    ManualPlanActive := FALSE;
    ManualRequiresSafeHeight := FALSE;
    ManualTargetChanged := FALSE;
    ManualComplete := FALSE;
    ManualTargetError := FALSE;
    LastActiveAxis := 0;
    AutoSegmentReady := FALSE;
  END_IF;
ELSIF Cmd = 0 THEN
  ModeState := 0;
  Step := 0;
  ManualSafeHeight := FALSE;
  ManualPhase := 0;
  ManualPlanActive := FALSE;
  ManualRequiresSafeHeight := FALSE;
  ManualTargetChanged := FALSE;
  ManualComplete := FALSE;
  ManualTargetError := FALSE;
  LastActiveAxis := 0;
  AutoSegmentReady := FALSE;
ELSIF (Cmd = 1) AND (LastCmd <> 1) THEN
  IF ManualPermitted THEN
    ModeState := 1;
    Step := 1;
    LastActiveAxis := 0;
    AutoSegmentReady := FALSE;
  ELSE
    Fault := 1;
  END_IF;
ELSIF Cmd = 4 THEN
  ManualValid := (ManualTarget1 >= -171.0) AND (ManualTarget1 <= 171.0)
                 AND (ManualTarget2 >= 130.0) AND (ManualTarget2 <= 360.0)
                 AND (ManualTarget3 >= 0.0) AND (ManualTarget3 <= 180.0)
                 AND (ManualTarget4 >= 12.0) AND (ManualTarget4 <= 70.0);
  ManualTargetError := NOT ManualValid;
  IF ManualPermitted AND ManualValid THEN
    IF (LastCmd <> 4)
       OR (ABS(ManualTarget1 - Captured1) > 0.01)
       OR (ABS(ManualTarget2 - Captured2) > 0.01)
       OR (ABS(ManualTarget3 - Captured3) > 0.01)
       OR (ABS(ManualTarget4 - Captured4) > 0.01) THEN
      ModeState := 4;
      Step := 0;
      Captured1 := ManualTarget1;
      Captured2 := ManualTarget2;
      Captured3 := ManualTarget3;
      Captured4 := ManualTarget4;
      ManualTargetChanged := TRUE;
      ManualPlanActive := TRUE;
      ManualComplete := FALSE;
      ManualRequiresSafeHeight := (ManualTarget2 < 280.0)
                                  AND ((ABS(Current1 - ManualTarget1) > 1.0)
                                       OR (ABS(Current3 - ManualTarget3) > 2.0));
      ManualSafeHeight := ManualRequiresSafeHeight;
      ManualPhase := 1;
      ManualAxisTarget2 := ManualTarget2;
      LastActiveAxis := 0;
    END_IF;
  ELSE
    Fault := 4;
  END_IF;
ELSIF (Cmd = 3) AND (LastCmd <> 3) THEN
  IF ManualPermitted AND (JogAxis >= 1) AND (JogAxis <= 4)
     AND ((JogDirection = -1) OR (JogDirection = 1)) THEN
    ModeState := 3;
    Step := 0;
    LastActiveAxis := 0;
  ELSE
    Fault := 7;
  END_IF;
END_IF;
LastCmd := Cmd;

IF ModeState = 1 THEN
  Permitted := AutoPermitted;
ELSE
  Permitted := ManualPermitted;
END_IF;

IF ((ModeState <> 0) AND (ModeState <> 1) AND NOT ManualPermitted)
   OR ((ModeState = 1) AND NOT ManualPermitted) THEN
  Fault := 1;
  ModeState := 0;
  Step := 0;
  ManualPhase := 0;
  ManualPlanActive := FALSE;
  ManualComplete := FALSE;
  LastActiveAxis := 0;
  AutoSegmentReady := FALSE;
END_IF;

IF ModeState = 1 THEN
  IF Step = 1 THEN
    DemoTarget1 := -68.754936; DemoTarget2 := 300.0; DemoTarget3 := 180.0; DemoTarget4 := 60.0;
  ELSIF Step = 2 THEN
    DemoTarget1 := -68.754936; DemoTarget2 := 150.0; DemoTarget3 := 180.0; DemoTarget4 := 60.0;
  ELSIF Step = 3 THEN
    DemoTarget1 := -68.754936; DemoTarget2 := 150.0; DemoTarget3 := 180.0; DemoTarget4 := 25.0;
  ELSIF Step = 4 THEN
    DemoTarget1 := -68.754936; DemoTarget2 := 320.0; DemoTarget3 := 180.0; DemoTarget4 := 25.0;
  ELSIF Step = 5 THEN
    DemoTarget1 := 80.214088; DemoTarget2 := 320.0; DemoTarget3 := 0.0; DemoTarget4 := 25.0;
  ELSIF Step = 6 THEN
    DemoTarget1 := 80.214088; DemoTarget2 := 180.0; DemoTarget3 := 0.0; DemoTarget4 := 25.0;
  ELSIF Step = 7 THEN
    DemoTarget1 := 80.214088; DemoTarget2 := 180.0; DemoTarget3 := 0.0; DemoTarget4 := 60.0;
  ELSIF Step = 8 THEN
    DemoTarget1 := 80.214088; DemoTarget2 := 300.0; DemoTarget3 := 0.0; DemoTarget4 := 60.0;
  ELSIF Step = 9 THEN
    DemoTarget1 := 80.214088; DemoTarget2 := 180.0; DemoTarget3 := 0.0; DemoTarget4 := 60.0;
  ELSIF Step = 10 THEN
    DemoTarget1 := 80.214088; DemoTarget2 := 180.0; DemoTarget3 := 0.0; DemoTarget4 := 25.0;
  ELSIF Step = 11 THEN
    DemoTarget1 := 80.214088; DemoTarget2 := 320.0; DemoTarget3 := 0.0; DemoTarget4 := 25.0;
  ELSIF Step = 12 THEN
    DemoTarget1 := -68.754936; DemoTarget2 := 320.0; DemoTarget3 := 180.0; DemoTarget4 := 25.0;
  ELSIF Step = 13 THEN
    DemoTarget1 := -68.754936; DemoTarget2 := 150.0; DemoTarget3 := 180.0; DemoTarget4 := 25.0;
  ELSIF Step = 14 THEN
    DemoTarget1 := -68.754936; DemoTarget2 := 150.0; DemoTarget3 := 180.0; DemoTarget4 := 60.0;
  ELSIF Step = 15 THEN
    DemoTarget1 := -68.754936; DemoTarget2 := 300.0; DemoTarget3 := 180.0; DemoTarget4 := 60.0;
  ELSE
    DemoTarget1 := 0.0; DemoTarget2 := 300.0; DemoTarget3 := 60.0; DemoTarget4 := 50.0;
  END_IF;
ELSIF ModeState = 2 THEN
  DemoTarget1 := 0.0; DemoTarget2 := 300.0; DemoTarget3 := 60.0; DemoTarget4 := 50.0;
ELSIF ModeState = 4 THEN
  DemoTarget1 := Captured1; DemoTarget2 := Captured2; DemoTarget3 := Captured3; DemoTarget4 := Captured4;
ELSE
  DemoTarget1 := Current1; DemoTarget2 := Current2; DemoTarget3 := Current3; DemoTarget4 := Current4;
END_IF;

Target1 := DemoTarget1;
Target2 := DemoTarget2;
Target3 := DemoTarget3;
Target4 := DemoTarget4;

AxisTarget2 := DemoTarget2;
ManualBaseReady := FALSE;
ManualExtensionReady := FALSE;
ManualSafeHeightReady := FALSE;
ManualHeightReady := FALSE;
ManualGripperReady := FALSE;

IF ModeState = 4 THEN
  ManualBaseReady := ABS(Current1 - Captured1) <= 1.0;
  ManualExtensionReady := ABS(Current3 - Captured3) <= 2.0;
  ManualHeightReady := ABS(Current2 - Captured2) <= 2.0;
  ManualGripperReady := ABS(Current4 - Captured4) <= 2.0;

  IF ManualTargetChanged THEN
    ManualTargetChanged := FALSE;
  END_IF;

  IF NOT ManualPlanActive THEN
    ManualPlanActive := TRUE;
    ManualComplete := FALSE;
    ManualPhase := 1;
    ManualRequiresSafeHeight := (Captured2 < 280.0)
                                AND (NOT ManualBaseReady OR NOT ManualExtensionReady);
    ManualSafeHeight := ManualRequiresSafeHeight;
    LastActiveAxis := 0;
  END_IF;

  IF ManualPhase = 0 THEN
    ManualPhase := 1;
    ManualComplete := FALSE;
    LastActiveAxis := 0;
  END_IF;

  IF ManualPhase = 1 THEN
    IF ManualRequiresSafeHeight THEN
      ManualAxisTarget2 := 300.0;
    ELSE
      ManualAxisTarget2 := Captured2;
    END_IF;
    AxisTarget2 := ManualAxisTarget2;

    IF ABS(Current2 - ManualAxisTarget2) <= 2.0 THEN
      ManualSafeHeightReady := TRUE;
      ManualPhase := 2;
      LastActiveAxis := 0;
    END_IF;
  END_IF;

  IF ManualPhase = 2 THEN
    IF ManualBaseReady THEN
      ManualPhase := 3;
      LastActiveAxis := 0;
    END_IF;
  END_IF;

  IF ManualPhase = 3 THEN
    IF ManualExtensionReady THEN
      IF ManualRequiresSafeHeight THEN
        ManualPhase := 4;
      ELSE
        ManualPhase := 5;
      END_IF;
      LastActiveAxis := 0;
    END_IF;
  END_IF;

  IF ManualPhase = 4 THEN
    ManualAxisTarget2 := Captured2;
    AxisTarget2 := ManualAxisTarget2;
    IF ManualHeightReady THEN
      ManualPhase := 5;
      LastActiveAxis := 0;
    END_IF;
  END_IF;

  IF ManualPhase = 5 THEN
    IF ManualGripperReady THEN
      ManualPhase := 6;
      ManualComplete := TRUE;
      LastActiveAxis := 0;
    END_IF;
  END_IF;

  IF ManualPhase = 6 THEN
    AxisTarget2 := Captured2;
    ManualComplete := ManualBaseReady AND ManualExtensionReady
                      AND ManualHeightReady AND ManualGripperReady;
  END_IF;

  IF ManualPhase = 1 THEN
    AxisTarget2 := ManualAxisTarget2;
    IF ABS(Current2 - ManualAxisTarget2) > 2.0 THEN ActiveAxis := 2; END_IF;
  ELSIF ManualPhase = 2 THEN
    IF NOT ManualBaseReady THEN ActiveAxis := 1; END_IF;
  ELSIF ManualPhase = 3 THEN
    IF NOT ManualExtensionReady THEN ActiveAxis := 3; END_IF;
  ELSIF ManualPhase = 4 THEN
    AxisTarget2 := Captured2;
    IF NOT ManualHeightReady THEN ActiveAxis := 2; END_IF;
  ELSIF ManualPhase = 5 THEN
    IF NOT ManualGripperReady THEN ActiveAxis := 4; END_IF;
  ELSE
    ActiveAxis := 0;
  END_IF;

  AtTarget := (ManualPhase = 6) AND ManualComplete
              AND ManualBaseReady AND ManualExtensionReady
              AND ManualHeightReady AND ManualGripperReady;
  ActiveStep := ManualPhase;
ELSIF ModeState = 2 THEN
  IF ABS(Current2 - AxisTarget2) > 2.0 THEN
    ActiveAxis := 2;
  ELSIF ABS(Current1 - DemoTarget1) > 1.0 THEN
    IF (Current2 >= 280.0) AND (DemoTarget2 >= 280.0) THEN ActiveAxis := 1; END_IF;
  ELSIF ABS(Current3 - DemoTarget3) > 2.0 THEN
    IF (Current2 >= 280.0) AND (DemoTarget2 >= 280.0) THEN ActiveAxis := 3; END_IF;
  ELSIF ABS(Current4 - DemoTarget4) > 2.0 THEN
    IF (ABS(Current1 - DemoTarget1) <= 1.0) AND (ABS(Current2 - DemoTarget2) <= 2.0)
       AND (ABS(Current3 - DemoTarget3) <= 2.0) THEN ActiveAxis := 4; END_IF;
  END_IF;
  AtTarget := (ActiveAxis = 0) AND (ABS(Current1 - DemoTarget1) <= 1.0)
              AND (ABS(Current2 - DemoTarget2) <= 2.0)
              AND (ABS(Current3 - DemoTarget3) <= 2.0)
              AND (ABS(Current4 - DemoTarget4) <= 2.0);
END_IF;

IF ModeState <> 1 THEN
  AutoSegmentReady := FALSE;
ELSIF NOT Permitted THEN
  AutoSegmentReady := FALSE;
ELSIF NOT AutoSegmentReady THEN
  AutoSegmentStart1 := Current1;
  AutoSegmentStart2 := Current2;
  AutoSegmentStart3 := Current3;
  AutoSegmentStart4 := Current4;
  AutoSegmentReady := TRUE;
END_IF;

AutoSegmentRunning := (ModeState = 1) AND Permitted AND AutoSegmentReady AND (Fault = 0);
AutoSegmentTimerA(IN := AutoSegmentRunning AND ((Step AND 1) <> 0), PT := T#1100ms);
AutoSegmentTimerB(IN := AutoSegmentRunning AND ((Step AND 1) = 0), PT := T#1100ms);
AutoSegmentDone := FALSE;

IF AutoSegmentRunning THEN
  IF (Step AND 1) <> 0 THEN
    P := TIME_TO_DINT(AutoSegmentTimerA.ET) / DINT_TO_REAL(1100);
    AutoSegmentDone := AutoSegmentTimerA.Q;
  ELSE
    P := TIME_TO_DINT(AutoSegmentTimerB.ET) / DINT_TO_REAL(1100);
    AutoSegmentDone := AutoSegmentTimerB.Q;
  END_IF;
  IF P < 0.0 THEN P := 0.0; END_IF;
  IF P > 1.0 THEN P := 1.0; END_IF;
  P := P * P * (3.0 - (2.0 * P));
  Current1 := AutoSegmentStart1 + ((DemoTarget1 - AutoSegmentStart1) * P);
  Current2 := AutoSegmentStart2 + ((DemoTarget2 - AutoSegmentStart2) * P);
  Current3 := AutoSegmentStart3 + ((DemoTarget3 - AutoSegmentStart3) * P);
  Current4 := AutoSegmentStart4 + ((DemoTarget4 - AutoSegmentStart4) * P);
  AnyMoving := TRUE;
  IF AutoSegmentDone THEN
    Current1 := DemoTarget1;
    Current2 := DemoTarget2;
    Current3 := DemoTarget3;
    Current4 := DemoTarget4;
    DonePulse := TRUE;
    Done := 1;
    DoneCounter := DoneCounter + 1;
    IF Step < 16 THEN
      Step := Step + 1;
    ELSE
      Step := 1;
    END_IF;
    AutoSegmentReady := FALSE;
  END_IF;
END_IF;

IF ActiveAxis = 1 THEN
  SegmentDurationMs := 1800;
ELSIF ActiveAxis = 2 THEN
  SegmentDurationMs := 2200;
ELSIF ActiveAxis = 3 THEN
  SegmentDurationMs := 1800;
ELSIF ActiveAxis = 4 THEN
  SegmentDurationMs := 1200;
ELSE
  SegmentDurationMs := 1800;
END_IF;

SegmentRunning := (ActiveAxis <> 0) AND (ActiveAxis = LastActiveAxis) AND (Fault = 0) AND Permitted;
IF ActiveAxis = 1 THEN
  SegmentTimer(IN := SegmentRunning, PT := T#1800ms);
ELSIF ActiveAxis = 2 THEN
  SegmentTimer(IN := SegmentRunning, PT := T#2200ms);
ELSIF ActiveAxis = 3 THEN
  SegmentTimer(IN := SegmentRunning, PT := T#1800ms);
ELSIF ActiveAxis = 4 THEN
  SegmentTimer(IN := SegmentRunning, PT := T#1200ms);
ELSE
  SegmentTimer(IN := FALSE, PT := T#1800ms);
END_IF;
IF ActiveAxis <> LastActiveAxis THEN
  IF ActiveAxis = 1 THEN SegmentStart1 := Current1; END_IF;
  IF ActiveAxis = 2 THEN SegmentStart2 := Current2; END_IF;
  IF ActiveAxis = 3 THEN SegmentStart3 := Current3; END_IF;
  IF ActiveAxis = 4 THEN SegmentStart4 := Current4; END_IF;
  LastActiveAxis := ActiveAxis;
ELSIF ActiveAxis <> 0 AND SegmentRunning THEN
  P := TIME_TO_DINT(SegmentTimer.ET) / DINT_TO_REAL(SegmentDurationMs);
  IF P < 0.0 THEN P := 0.0; END_IF;
  IF P > 1.0 THEN P := 1.0; END_IF;
  P := P * P * (3.0 - (2.0 * P));
  IF ActiveAxis = 1 THEN Current1 := SegmentStart1 + ((DemoTarget1 - SegmentStart1) * P); END_IF;
  IF ActiveAxis = 2 THEN Current2 := SegmentStart2 + ((AxisTarget2 - SegmentStart2) * P); END_IF;
  IF ActiveAxis = 3 THEN Current3 := SegmentStart3 + ((DemoTarget3 - SegmentStart3) * P); END_IF;
  IF ActiveAxis = 4 THEN Current4 := SegmentStart4 + ((DemoTarget4 - SegmentStart4) * P); END_IF;
  AnyMoving := TRUE;
END_IF;

JogPulseTimer(IN := (ModeState = 3) AND (Cmd = 3) AND (JogEnable <> 0)
                    AND Permitted AND NOT JogPulseTimer.Q, PT := T#50ms);
IF (ModeState = 3) AND (Cmd = 3) AND (JogEnable <> 0) AND Permitted AND JogPulseTimer.Q THEN
  IF JogAxis = 1 THEN
    Current1 := Current1 + (INT_TO_REAL(JogDirection) * 1.5);
    IF Current1 < -171.0 THEN Current1 := -171.0; END_IF;
    IF Current1 > 171.0 THEN Current1 := 171.0; END_IF;
  ELSIF JogAxis = 2 THEN
    Current2 := Current2 + (INT_TO_REAL(JogDirection) * 4.0);
    IF Current2 < 130.0 THEN Current2 := 130.0; END_IF;
    IF Current2 > 360.0 THEN Current2 := 360.0; END_IF;
  ELSIF JogAxis = 3 THEN
    IF Current2 >= 280.0 THEN
      Current3 := Current3 + (INT_TO_REAL(JogDirection) * 4.0);
      IF Current3 < 0.0 THEN Current3 := 0.0; END_IF;
      IF Current3 > 180.0 THEN Current3 := 180.0; END_IF;
    END_IF;
  ELSIF JogAxis = 4 THEN
    IF (ABS(Current1 - DemoTarget1) <= 1.0) AND (ABS(Current2 - DemoTarget2) <= 2.0)
       AND (ABS(Current3 - DemoTarget3) <= 2.0) THEN
      Current4 := Current4 + (INT_TO_REAL(JogDirection) * 2.0);
      IF Current4 < 12.0 THEN Current4 := 12.0; END_IF;
      IF Current4 > 70.0 THEN Current4 := 70.0; END_IF;
    END_IF;
  END_IF;
  AnyMoving := TRUE;
END_IF;

SettleTimer(IN := ((ModeState = 2) OR (ModeState = 4))
                   AND AtTarget AND Permitted AND (Fault = 0), PT := T#200ms);
IF SettleTimer.Q AND (Fault = 0) THEN
  DonePulse := TRUE;
  Done := 1;
  DoneCounter := DoneCounter + 1;
  ModeState := 0;
  Step := 0;
  LastActiveAxis := 0;
END_IF;

IF Fault <> 0 THEN
  ModeState := 0;
  Step := 0;
  LastActiveAxis := 0;
  AutoSegmentReady := FALSE;
END_IF;

IF Fault <> 0 THEN
  Status := 3;
ELSIF DonePulse THEN
  Status := 2;
ELSIF (ModeState = 1) AND NOT Permitted THEN
  Status := 0;
ELSIF (ModeState <> 0) AND Permitted AND (AnyMoving OR (ActiveAxis <> 0)) THEN
  Status := 1;
ELSE
  Status := 0;
END_IF;

IF ModeState = 1 THEN
  ActiveMode := 1;
ELSIF ModeState = 3 THEN
  ActiveMode := 3;
ELSIF (ModeState = 4) OR (ModeState = 2) THEN
  ActiveMode := 4;
ELSE
  ActiveMode := 0;
END_IF;
IF ModeState = 4 THEN
  ActiveStep := ManualPhase;
ELSE
  ActiveStep := Step;
END_IF;
AlarmCode := Fault;

RunMask := 0;
DirectionMask := 0;
CmdQ1toQ8Mask := 0;
IF (ModeState = 1) AND Permitted AND (Fault = 0) THEN
  IF ABS(DemoTarget1 - Current1) > 0.01 THEN RunMask := RunMask OR 1; END_IF;
  IF ABS(DemoTarget2 - Current2) > 0.01 THEN RunMask := RunMask OR 2; END_IF;
  IF ABS(DemoTarget3 - Current3) > 0.01 THEN RunMask := RunMask OR 4; END_IF;
  IF ABS(DemoTarget4 - Current4) > 0.01 THEN RunMask := RunMask OR 8; END_IF;
  IF ((RunMask AND 1) <> 0) AND (DemoTarget1 >= Current1) THEN DirectionMask := DirectionMask OR 1; END_IF;
  IF ((RunMask AND 2) <> 0) AND (DemoTarget2 >= Current2) THEN DirectionMask := DirectionMask OR 2; END_IF;
  IF ((RunMask AND 4) <> 0) AND (DemoTarget3 >= Current3) THEN DirectionMask := DirectionMask OR 4; END_IF;
  IF ((RunMask AND 8) <> 0) AND (DemoTarget4 >= Current4) THEN DirectionMask := DirectionMask OR 8; END_IF;
ELSIF (ModeState <> 0) AND Permitted AND (Fault = 0) AND (ActiveAxis <> 0) THEN
  IF ActiveAxis = 1 THEN RunMask := 1;
  ELSIF ActiveAxis = 2 THEN RunMask := 2;
  ELSIF ActiveAxis = 3 THEN RunMask := 4;
  ELSIF ActiveAxis = 4 THEN RunMask := 8;
  END_IF;
  IF ActiveAxis = 1 THEN
    IF DemoTarget1 >= Current1 THEN DirectionMask := 1; END_IF;
  ELSIF ActiveAxis = 2 THEN
    IF DemoTarget2 >= Current2 THEN DirectionMask := 2; END_IF;
  ELSIF ActiveAxis = 3 THEN
    IF DemoTarget3 >= Current3 THEN DirectionMask := 4; END_IF;
  ELSIF ActiveAxis = 4 THEN
    IF DemoTarget4 >= Current4 THEN DirectionMask := 8; END_IF;
  END_IF;
END_IF;

IF (RunMask AND 1) <> 0 THEN CmdQ1toQ8Mask := CmdQ1toQ8Mask OR 3; END_IF;
IF (RunMask AND 2) <> 0 THEN CmdQ1toQ8Mask := CmdQ1toQ8Mask OR 12; END_IF;
IF (RunMask AND 4) <> 0 THEN CmdQ1toQ8Mask := CmdQ1toQ8Mask OR 48; END_IF;
IF (RunMask AND 8) <> 0 THEN CmdQ1toQ8Mask := CmdQ1toQ8Mask OR 192; END_IF;

Pos1 := Current1;
Pos2 := Current2;
Pos3 := Current3;
Pos4 := Current4;

IF ModeState = 0 THEN
  Target1 := Current1;
  Target2 := Current2;
  Target3 := Current3;
  Target4 := Current4;
END_IF;

RealBits := ADR(Pos1);
Pos1High := TO_UINT(SHR(RealBits^, 16));
Pos1Low := TO_UINT(RealBits^ AND 16#0000FFFF);
RealBits := ADR(Pos2);
Pos2High := TO_UINT(SHR(RealBits^, 16));
Pos2Low := TO_UINT(RealBits^ AND 16#0000FFFF);
RealBits := ADR(Pos3);
Pos3High := TO_UINT(SHR(RealBits^, 16));
Pos3Low := TO_UINT(RealBits^ AND 16#0000FFFF);
RealBits := ADR(Pos4);
Pos4High := TO_UINT(SHR(RealBits^, 16));
Pos4Low := TO_UINT(RealBits^ AND 16#0000FFFF);
RealBits := ADR(Target1);
Target1High := TO_UINT(SHR(RealBits^, 16));
Target1Low := TO_UINT(RealBits^ AND 16#0000FFFF);
RealBits := ADR(Target2);
Target2High := TO_UINT(SHR(RealBits^, 16));
Target2Low := TO_UINT(RealBits^ AND 16#0000FFFF);
RealBits := ADR(Target3);
Target3High := TO_UINT(SHR(RealBits^, 16));
Target3Low := TO_UINT(RealBits^ AND 16#0000FFFF);
RealBits := ADR(Target4);
Target4High := TO_UINT(SHR(RealBits^, 16));
Target4Low := TO_UINT(RealBits^ AND 16#0000FFFF);

(* ---- watertank.st ---- *)
  VAR
    openOutletValve : BOOL AT %QX0.1;
    openInletValve : BOOL AT %QX0.4;
    outletValveOpenStatus : BOOL AT %QX0.3;
    inletValveOpenStatus : BOOL AT %QX0.5;
    airValveOpenStatus : BOOL AT %QX0.6;
    level : INT AT %IW2;
    level_max : INT AT %IW3;
    level_min : INT := 10;
  END_VAR

IF (level >= level_max) AND airValveOpenStatus THEN
  openOutletValve := TRUE;
  outletValveOpenStatus := TRUE;
  openInletValve := FALSE;
  inletValveOpenStatus := FALSE;
END_IF;

IF (level < (level_max - level_min)) AND airValveOpenStatus THEN
  openOutletValve := FALSE;
  outletValveOpenStatus := FALSE;
  openInletValve := TRUE;
  inletValveOpenStatus := TRUE;
END_IF;

IF NOT airValveOpenStatus THEN
  openOutletValve := FALSE;
  outletValveOpenStatus := FALSE;
  openInletValve := FALSE;
  inletValveOpenStatus := FALSE;
END_IF;
